// TIA Portal V20 export
// export: Created 2026-10-20T18:54:27.5257907Z, ExportSetting None, DisplayName Totally Integrated Automation Portal, DisplayVersion V20 Update 6, DisplayName TIA Portal Openness, DisplayVersion V20 Update 6, DisplayName TIA Portal Version Control Interface, DisplayVersion V20 Update 6, DisplayName SINAMICS Startdrive Advanced, DisplayVersion V20 SP1, DisplayName SINAMICS Startdrive G130, G150, S120, S150, SINAMICS MV, G220, S200, S210, DisplayVersion V20 SP1, DisplayName SINAMICS Startdrive G110M, G120, G120C, G120D, G120P, G115D, DisplayVersion V20 SP1, DisplayName STEP 7 Professional, DisplayVersion V20 Update 6, DisplayName STEP 7 Safety, DisplayVersion V20 Update 2, DisplayName WinCC Basic/Comfort/Advanced, DisplayVersion V20 Update 6, DisplayName WinCC Unified, DisplayVersion V20 Update 6
VAR_GLOBAL   // PLC tag table "VTD_HMI"
   Start_InBarcodeStation_HMI AT %M25.4 : Bool;
   VTD_Move_To_Level_HMI AT %MW1006 : UInt;
   VTD_Mode_Change_HMI AT %MW1000 : UInt;
   VTD_Manual_Down_HMI AT %M3.4 : Bool;
   VTD_Start_Teach_HMIs AT %M4.4 : Bool;
   VTD_Pallet_Type_HMI AT %MW1002 : UInt;
   VTD_Manual_Up_HMI AT %M3.3 : Bool;
   VTD_Task_ID_HMI AT %MW1004 : UInt;
   VTD_Reset_HMIs AT %M2.5 : Bool;
   VTD_Enable_HMI AT %M2.4 : Bool;
   VTD_Progress_HMI AT %MW1040 : Int;
   VTD_Stop_HMI AT %M3.2 : Bool;
   VTD_Manual_LP_Extend_HMIs AT %M4.3 : Bool;
   VTD_Manual_LP_Retract_HMIs AT %M3.5 : Bool;
   VTD_ID_HMI AT %MW12 : UInt;
   VTD_Cnv_Occupied AT %M25.6 : Bool;
   VTD_Motor_Status_HMI AT %MW120 : UInt;
   VTD_ID_HMI_OLD AT %MW116 : UInt;
   VTD_LE_Error_HMI AT %M1024.0 : Bool;
   VTD_Mode_HMI AT %MW1008 : UInt;
   VTD_Encoder_Delta_HMI AT %MD1028 : Real;
   VTD_Warning_HMI AT %M11.1 : Bool;
   VTD_Current_Level_HMI AT %MW1014 : UInt;
   VTD_Error_HMI AT %M11.0 : Bool;
   VTD_Current_Task_ID_HMI AT %MW1012 : UInt;
   VTD_Pallet_Loaded_HMI AT %MW1018 : UInt;
   VTD_Stopped_HMI AT %M11.3 : Bool;
   VTD_SM_State_HMI AT %MW1022 : UInt;
   VTD_Shuttle_Loaded_HMI AT %MW1020 : UInt;
   VTD_LP_State_HMI AT %MW1016 : UInt;
   VTD_AE_HMI AT %MD1032 : Real;
   VTD_Docked_HMI AT %M11.5 : Bool;
   VTD_AE_Error_HMI AT %M1026.0 : Bool;
   VTD_Enabled_HMI AT %M11.2 : Bool;
   VTD_Current_Task_Type_HMI AT %MW1010 : UInt;
   VTD_Running_HMI AT %M11.4 : Bool;
   VTD_LE_HMI AT %MD1143 : Real;
   VTD_Motor_Actual_Speed_HMI AT %MW134 : UInt;
   VTD_Motor_SetPoint_HMI AT %MW132 : UInt;
   VTD_Motor_Actual_Current_HMI AT %MD128 : Real;
   VTD_Motor_Ready_HMI AT %M136.1 : Bool;
   "Chain Slack 1" AT %M102.0 : Bool;
   "Chain Slack 3" AT %M104.1 : Bool;
   "Chain Slack 2" AT %M104.0 : Bool;
   "Chain Slack 4" AT %M104.2 : Bool;
   VTD_LE_Speed_HMI AT %MW118 : Int;
   "BCD_Disable_Trigger_HMI(5)" AT %M26.4 : Bool;
   "BCD_Enable_Trigger_HMI(3)" AT %M25.0 : Bool;
   "BCD_Disable_Trigger_HMI(4)" AT %M26.3 : Bool;
   "BCD_Disable_Trigger_HMI(3)" AT %M26.2 : Bool;
   "BCD_Test_Comm_HMI(5)" AT %M14.6 : Bool;
   "BCD_Disable_Trigger_HMI(2)" AT %M26.1 : Bool;
   "BCD_Test_Comm_HMI(2)" AT %M14.3 : Bool;
   "BCD_Test_Comm_HMI(4)" AT %M14.5 : Bool;
   "BCD_Test_Comm_HMI(1)" AT %M14.0 : Bool;
   "BCD_Test_Comm_HMI(3)" AT %M14.4 : Bool;
   "BCD_Enable_Trigger_HMI(4)" AT %M25.7 : Bool;
   "BCD_Enable_Trigger_HMI(5)" AT %M26.0 : Bool;
   "BCD_Enable_Trigger_HMI(2)" AT %M14.7 : Bool;
   "BCD_Enable_Trigger_HMI(1)" AT %M14.1 : Bool;
   "BCD_Disable_Trigger_HMI(1)" AT %M14.2 : Bool;
   Safety_OK_HMI AT %M26.5 : Bool;
   VTD_Moving_To_Level AT %MW160 : UInt;
   VTD_Speed_mm_s AT %MD166 : Real;
   VTD_Level_Below_Extractor AT %MW164 : UInt;
   VTD_Actual_Torque AT %MW176 : UInt;
END_VAR
